(* IEC 61131-3 sources: plc-process-lib/tools/demo/src/POUs/F_DemoInterp, 2 files *)

(* ---- F_DemoInterp.decl.st ---- *)
// Назначение: линейная интерполяция между двумя точками профиля сценария (время, значение).
//             Вне отрезка — значение ближайшего конца; отрезок нулевой длины — конечное значение.
// Автор:      kr0nsch
// Версия:     0.1.0
// Документ:   docs/media/data/ (профили сценариев); tools/demo/README.md
FUNCTION F_DemoInterp : REAL
VAR_INPUT
    lrT0_s : LREAL;   // начало отрезка, с
    rV0    : REAL;    // значение в начале
    lrT1_s : LREAL;   // конец отрезка, с
    rV1    : REAL;    // значение в конце
    lrT_s  : LREAL;   // момент, с
END_VAR

(* ---- F_DemoInterp.impl.st ---- *)
IF lrT_s <= lrT0_s THEN
    F_DemoInterp := rV0;
ELSIF lrT_s >= lrT1_s OR lrT1_s <= lrT0_s THEN
    F_DemoInterp := rV1;
ELSE
    F_DemoInterp := LREAL_TO_REAL(REAL_TO_LREAL(rV0)
                    + REAL_TO_LREAL(rV1 - rV0) * (lrT_s - lrT0_s) / (lrT1_s - lrT0_s));
END_IF
